TYPE ST_MCExecuteParam :
STRUCT
	fTargetVelocity: LREAL;
	eCommand: E_Command;
	ePlanningMode: E_PlanningMode;
	stStartPosition: ST_Point;
	stEndPosition: ST_Point;
END_STRUCT
END_TYPE

(* stored: Version 1.1.0.1, ProductVersion 3.1.4024.12
   DUT ST_MCExecuteParam: Id {2b529d63-564a-4910-99fa-386a1f0fd1b2} *)
